(* Communication structure from plc to drive *)

TYPE ST_PLCTOFORCE :
STRUCT

END_STRUCT
END_TYPE

(* stored: Version 1.1.0.1, ProductVersion 3.1.4024.15
   DUT ST_PLCTOFORCE: Id {383702f3-e446-4c74-9dff-ef06483bc061} *)
